(* Logix 5000 project; controller NWGG 1756-L72 rev 35.12; software revision 35.00; part 10 of 19 *)
(* tags used below, declared in another part *)
   _11_GATE_PO : ALIAS FOR I16[0];
   _123_COMPUW : ALIAS FOR I18[7];
   _12_GATE_PO : ALIAS FOR I16[1];
   _13_GATE_PO : ALIAS FOR I16[2];
   _14_GATE_PO : ALIAS FOR I16[3];
   _15_GATE_PO : ALIAS FOR I16[4];
   _16_GATE_PO : ALIAS FOR I16[5];
   _17_GATE_PO : ALIAS FOR I16[6];
   _21_GATE_PO : ALIAS FOR I16[7];
   _22_GATE_PO : ALIAS FOR I17[0];
   _23_GATE_PO : ALIAS FOR I17[1];
   _24_GATE_PO : ALIAS FOR I17[2];
   _25_GATE_PO : ALIAS FOR I17[3];
   _26_GATE_PO : ALIAS FOR I17[4];
   _27_GATE_PO : ALIAS FOR I17[5];
   _27_GATE_PO1 : ALIAS FOR N14[27];
   _28_GATE_PO : ALIAS FOR I17[6];
   _28_GATE_PO1 : ALIAS FOR N14[28];
   _29_GATE_PO : ALIAS FOR I17[7];
   _29_GATE_PO1 : ALIAS FOR N14[29];
   _41_GATE_PO : ALIAS FOR I18[0];
   _42_GATE_PO : ALIAS FOR I18[1];
   _701K_GATE2 : ALIAS FOR B21[11].2;
   _701K_VALVE : ALIAS FOR O13.10;
   Beta : BOOL;
   Calibration_Max : REAL;
   Cleaning_Motors : udt_Motor[100];
   cpTicketBinActive : DINT;
   cpTicketBinSet : DINT;
   Dev : DINT;
   I18 : INT[16];
   I18_002 : ALIAS FOR I18[2];
   I18_003 : ALIAS FOR I18[3];
   indexTbl : DINT;
   indexTRTTbl : DINT;
   InEUMax : REAL;
   MAIN_TIMER : ALIAS FOR T11[0];
   O11_000_Bit09 : ALIAS FOR O11.9;
   O11_000_Bit10 : ALIAS FOR O11.10;
   O11_000_Bit11 : ALIAS FOR O11.11;
   O11_000_Bit12 : ALIAS FOR O11.12;
   O11_000_Bit13 : ALIAS FOR O11.13;
   O11_000_Bit14 : ALIAS FOR O11.14;
   O12_000_Bit00 : ALIAS FOR O12.0;
   O12_000_Bit01 : ALIAS FOR O12.1;
   O12_000_Bit02 : ALIAS FOR O12.2;
   O16 : INT[12];
   O17 : INT[12];
   O18 : INT[12];
   O9_000_Bit00 : ALIAS FOR O9.0;
   SCREENINGS : ALIAS FOR I7.15;
   sendData : BOOL;
   sendData1 : BOOL;
   spBinGateRates : DINT[50];
   spCapGrossWt : BOOL;
   spCapTareWt : BOOL;
   spCreateTicket : BOOL;
   spShowCreateTicketPB : BOOL;
   spTicketBinActive : DINT;
   spTicketBinSet : DINT;
   spTicketProcessing : BOOL;
   spTicketProcessStr : BOOL;
   spTicketTableBay1GrsWt : DINT;
   spTicketTableBay1Wt : DINT;
   spVAR_BINARRAY : STRING[50];
   sqlIndex : DINT;
   sqlIndex1 : DINT;
   sqlNewTreatment : BOOL;
   sqlNewTreatments_ONS : DINT;
   sqlNewVariety : BOOL;
   sqlNewVariety_ONS : DINT;
   sqlTreatID : DINT;
   sqlTreatmentsRevd : DINT;
   sqlTreatRate : DINT;
   sqlTrtSendDelayTMR : TIMER;
   sqlVaritiesRevd : DINT;
   sqlVarityID : DINT;
   sqlVarityRate : DINT;
   sqlVarSendDelayTMR : TIMER;
   SWW_Index : DINT;
   SWW_Variety_DB : Varieties_DB[100];
   T11_AUTO_M : ALIAS FOR B3[11].1;
   T11_AUTO_S : ALIAS FOR B3[11].14;
   T11_SET_LO : ALIAS FOR B3[11].13;
   T12_AUTO_M : ALIAS FOR B3[12].1;
   T12_AUTO_S : ALIAS FOR B3[12].14;
   T12_SET_LO : ALIAS FOR B3[12].13;
   T13_AUTO_M : ALIAS FOR B3[13].1;
   T13_AUTO_S : ALIAS FOR B3[13].14;
   T13_SET_LO : ALIAS FOR B3[13].13;
   T14_AUTO_M : ALIAS FOR B3[14].1;
   T14_AUTO_S : ALIAS FOR B3[14].14;
   T14_SET_LO : ALIAS FOR B3[14].13;
   T15_AUTO_M : ALIAS FOR B3[15].1;
   T15_AUTO_S : ALIAS FOR B3[15].14;
   T15_SET_LO : ALIAS FOR B3[15].13;
   T16_AUTO_M : ALIAS FOR B3[16].1;
   T16_AUTO_S : ALIAS FOR B3[16].14;
   T16_SET_LO : ALIAS FOR B3[16].13;
   T17_AUTO_M : ALIAS FOR B3[17].1;
   T17_AUTO_S : ALIAS FOR B3[17].14;
   T17_SET_LO : ALIAS FOR B3[17].13;
   T21_AUTO_M : ALIAS FOR B3[21].1;
   T21_AUTO_S : ALIAS FOR B3[21].14;
   T21_SET_LO : ALIAS FOR B3[21].13;
   T22_AUTO_M : ALIAS FOR B3[22].1;
   T22_AUTO_S : ALIAS FOR B3[22].14;
   T22_SET_LO : ALIAS FOR B3[22].13;
   T23_AUTO_M : ALIAS FOR B3[23].1;
   T23_AUTO_S : ALIAS FOR B3[23].14;
   T23_SET_LO : ALIAS FOR B3[23].13;
   T24_AUTO_M : ALIAS FOR B3[24].1;
   T24_AUTO_S : ALIAS FOR B3[24].14;
   T24_SET_LO : ALIAS FOR B3[24].13;
   T25_AUTO_M : ALIAS FOR B3[25].1;
   T25_AUTO_S : ALIAS FOR B3[25].14;
   T25_SET_LO : ALIAS FOR B3[25].13;
   T26_AUTO_M : ALIAS FOR B3[26].1;
   T26_AUTO_S : ALIAS FOR B3[26].14;
   T26_SET_LO : ALIAS FOR B3[26].13;
   T27_AUTO_M : ALIAS FOR B3[27].1;
   T27_CLOSE1 : ALIAS FOR B3[27].9;
   T27_CLOSE2 : ALIAS FOR B3[27].11;
   T27_FAULT : ALIAS FOR B3[27].15;
   T27_GATE_C : ALIAS FOR C5[27];
   T27_HOLD_A : ALIAS FOR B3[27].3;
   T27_HOLD_M : ALIAS FOR B3[27].6;
   T27_OPEN_A : ALIAS FOR B3[27].8;
   T27_OPEN_M1 : ALIAS FOR B3[27].10;
   T27_RELEAS : ALIAS FOR B3[27].5;
   T27_RESET : ALIAS FOR B3[27].7;
   T27_SET_AU : ALIAS FOR B3[27].2;
   T27_STOP_A : ALIAS FOR B3[27].4;
   T28_AUTO_M : ALIAS FOR B3[28].1;
   T28_CLOSE1 : ALIAS FOR B3[28].9;
   T28_CLOSE2 : ALIAS FOR B3[28].11;
   T28_FAULT : ALIAS FOR B3[28].15;
   T28_GATE_C : ALIAS FOR C5[28];
   T28_HOLD_A : ALIAS FOR B3[28].3;
   T28_HOLD_M : ALIAS FOR B3[28].6;
   T28_OPEN_A : ALIAS FOR B3[28].8;
   T28_OPEN_M1 : ALIAS FOR B3[28].10;
   T28_RELEAS : ALIAS FOR B3[28].5;
   T28_RESET : ALIAS FOR B3[28].7;
   T28_SET_AU : ALIAS FOR B3[28].2;
   T28_STOP_A : ALIAS FOR B3[28].4;
   T29_AUTO_M : ALIAS FOR B3[29].1;
   T29_CLOSE1 : ALIAS FOR B3[29].9;
   T29_CLOSE2 : ALIAS FOR B3[29].11;
   T29_FAULT : ALIAS FOR B3[29].15;
   T29_GATE_C : ALIAS FOR C5[29];
   T29_HOLD_A : ALIAS FOR B3[29].3;
   T29_HOLD_M : ALIAS FOR B3[29].6;
   T29_OPEN_A : ALIAS FOR B3[29].8;
   T29_OPEN_M1 : ALIAS FOR B3[29].10;
   T29_RELEAS : ALIAS FOR B3[29].5;
   T29_RESET : ALIAS FOR B3[29].7;
   T29_SET_AU : ALIAS FOR B3[29].2;
   T29_STOP_A : ALIAS FOR B3[29].4;
   TestTag : REAL;
   TicketTreatPumpActive : DINT;
   TicketTreatPumpSet : DINT;
   tpCreateTicket : BOOL;
   tpCreateTicketRecvd : DINT;
   tpLocation : DINT;
   tpNewGrossWt : BOOL;
   tpNewGrossWtRecvd : DINT;
   tpNewGrossWtSent : BOOL;
   tpNewTareWt : BOOL;
   tpNewTareWtRecvd : DINT;
   tpNewTareWtSent : BOOL;
   tpShowGrossPB : BOOL;
   tpShowTarePB : BOOL;
   tpVarsTrtsComplete : BOOL;
   TRT_CNT : DINT;
   Trt_CntStore : DINT;
   TRT_TickettableItemNo : DINT[50];
   TRT_TICKETtableRate : DINT[100];
   VAR_CNT : DINT;
   VAR_CNT_ONS : DINT;
   Var_CntStore : DINT;
   VAR_TICKETtable : STRING[20];
   VAR_TickettableItemNo : DINT[50];
   VAR_TICKETtableRate : DINT[100];
   VarTrimTemp : STRING;
   zzztmpTANKtest : DINT[10];
   zzzzTestGrossWt : BOOL;
   zzzzTestTareWt : BOOL;
(* _2_MAIN, continued *)

ROUTINE _701_KValve   (* ladder *)
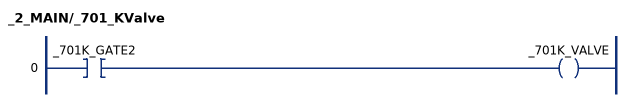
   0: XIC(_701K_GATE2)OTE(_701K_VALVE);
END_ROUTINE

ROUTINE _99_Scaling   (* function block diagram *)
   SHEET 1
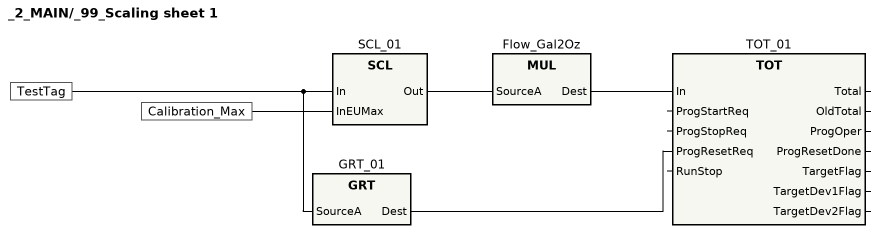
   GRT_01 : GRT(SourceA := TestTag);
   SCL_01 : SCL(In := TestTag, InEUMax := Calibration_Max);
   Flow_Gal2Oz : MUL(SourceA := SCL_01.Out);
   TOT_01 : TOT(In := Flow_Gal2Oz.Dest, ProgResetReq := GRT_01.Dest);   // unwired pins: ProgStartReq ProgStopReq Total OldTotal ProgOper RunStop ProgResetDone TargetFlag TargetDev1Flag TargetDev2Flag
   SHEET 2
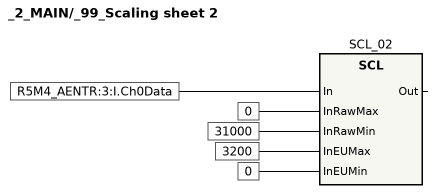
   SCL_02 : SCL(In := R5M4_AENTR:3:I.Ch0Data, InRawMax := 0, InRawMin := 31000, InEUMax := 3200, InEUMin := 0);   // unwired pins: Out
END_ROUTINE
END_PROGRAM

PROGRAM Amp_Guages   (* main routine Amp_Guages *)
VAR
   SCL_AMP_Belt11 : SCALE := (In := 28.19336, InRawMax := 6000.0, InEUMax := 1.61, Out := 0.007565218);
   SCL_AMP_Belt11_01 : SCALE := (In := 23.047852, InRawMax := 9000.0, InRawMin := 20.0, InEUMax := 2.15, Out := 0.0007297195);
   SCL_AMP_Belt11_02 : SCALE := (In := 4111.1504, InRawMax := 7000.0, InRawMin := 20.0, InEUMax := 1.61, Out := 0.94366074);
   SCL_AMP_Belt11_03 : SCALE := (In := 7592.727, InRawMax := 13000.0, InRawMin := 20.0, InEUMax := 3.88, Out := 2.2636504);
END_VAR

ROUTINE Amp_Guages   (* function block diagram *)
   SHEET 1
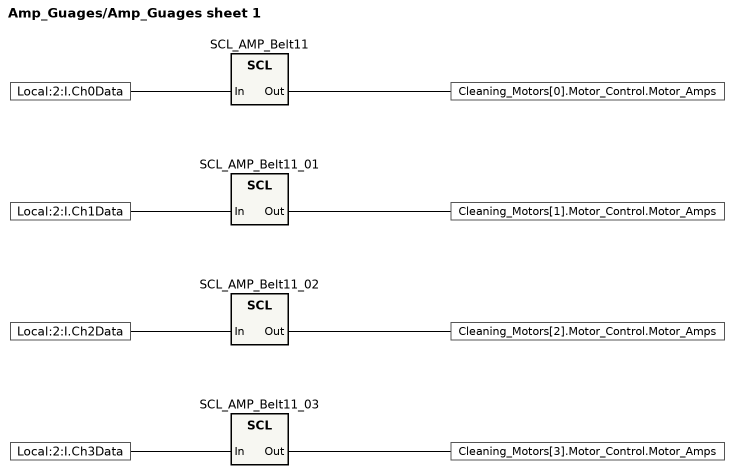
   SCL_AMP_Belt11 : SCL(In := Local:2:I.Ch0Data);
   SCL_AMP_Belt11_01 : SCL(In := Local:2:I.Ch1Data);
   SCL_AMP_Belt11_02 : SCL(In := Local:2:I.Ch2Data);
   SCL_AMP_Belt11_03 : SCL(In := Local:2:I.Ch3Data);
   Cleaning_Motors[0].Motor_Control.Motor_Amps := SCL_AMP_Belt11.Out;
   Cleaning_Motors[1].Motor_Control.Motor_Amps := SCL_AMP_Belt11_01.Out;
   Cleaning_Motors[2].Motor_Control.Motor_Amps := SCL_AMP_Belt11_02.Out;
   Cleaning_Motors[3].Motor_Control.Motor_Amps := SCL_AMP_Belt11_03.Out;
END_ROUTINE
END_PROGRAM

PROGRAM Load_Requests   (* main routine Main *)

ROUTINE Main   (* ladder *)
END_ROUTINE
END_PROGRAM

PROGRAM Main   (* main routine Main *)
VAR
   alm_Development : ALARM_DIGITAL;
   Beta_Mode : BOOL;
END_VAR

ROUTINE Main   (* ladder *)
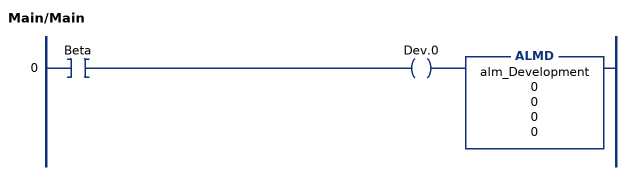
   0: XIC(Beta)OTE(Dev.0)ALMD(alm_Development,0,0,0,0);
END_ROUTINE
END_PROGRAM

PROGRAM MainProgram   (* main routine MainRoutine *)
VAR
   Alm_Test : BOOL := 1;
   ATestAck : BOOL;
   ATestPDis : BOOL;
   ATestPEna : BOOL;
   ATestReset : BOOL;
   BIN13test : BOOL;
   CleaningBinVarieties : STRING[10] := ([2] := 'hale', [3] := 'Hale full', [4] := 'Hale', [6] := 'HD307 Screenings');
   CTR_Scale_Accum_Rate_Index : COUNTER;
   Flow_Gal2Oz : FBD_MATH := (SourceA := 4000.0, SourceB := 0.25, Dest := 1000.0);
   GRT_01 : FBD_COMPARE := (SourceB := 75.0);
   Rate_Tmr : TIMER := (PRE := 1000, ACC := 610, TT := 1, DN := 1);
   Scale_Avg_Ctr : COUNTER := (PRE := 10, ACC := 2, CU := 1);
   ScaleWeights : DINT[60];
   SCL_01 : SCALE := (InRawMax := 100.0, InEUMax := 4000.0);
   SCL_02 : SCALE := (In := 16384.0, InRawMax := 13975.0, InRawMin := 578.0, InEUMax := 3000.0, Limiting := 1, Out := 3000.0, MaxAlarm := 1);
   Tare : DINT;
   tmr_User_Cancel : TIMER := (PRE := 5000, ACC := 5004, EN := 1, DN := 1);
   tmrWeightTest : TIMER := (PRE := 500, ACC := 112, EN := 1, TT := 1);
   TOT_01 : TOTALIZER := (TimeBase := 1, Gain := 1.0, ProgProgReq := 1, ProgStartReq := 1, ProgStopReq := 1, RTSTime := 1, Total := 4074.4673, OldTotal := 9541.935, ProgOper := 1, TargetFlag := 1, TargetDev1Flag := 1, TargetDev2Flag := 1, LowInCutoffFlag := 1, DeltaT := 0.016);
   Truck_Scale_Control : Truck_Scale_Control[2];
   Weight_Seed : DINT := 10;
END_VAR

ROUTINE _100_VarCfg   (* ladder *)
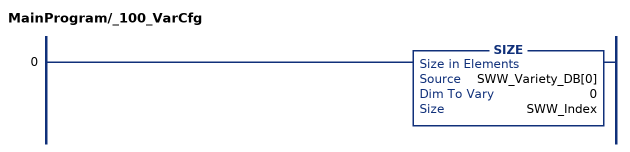
   0: SIZE(SWW_Variety_DB[0],0,SWW_Index);
END_ROUTINE

ROUTINE _31_TANK_27   (* ladder *)
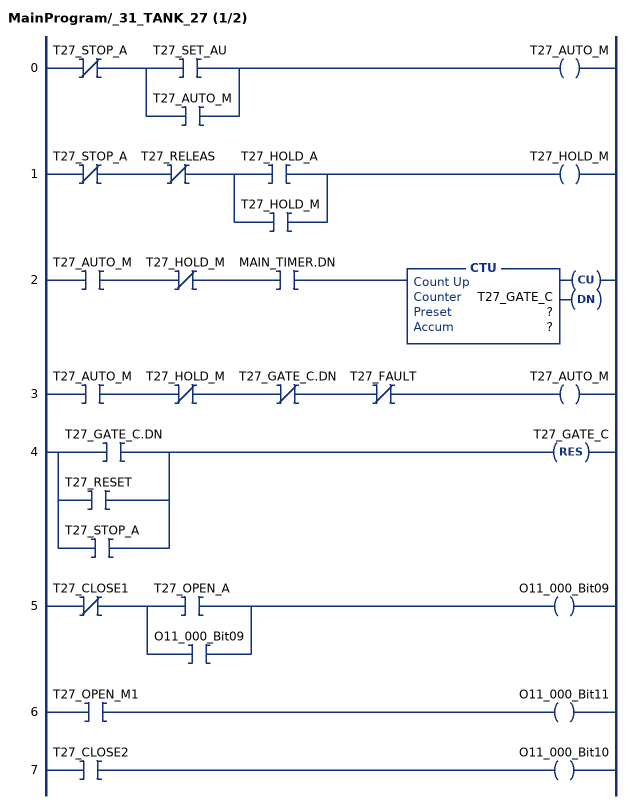
   0: XIO(T27_STOP_A)[XIC(T27_SET_AU) ,XIC(T27_AUTO_M) ]OTE(T27_AUTO_M);
   1: XIO(T27_STOP_A)XIO(T27_RELEAS)[XIC(T27_HOLD_A) ,XIC(T27_HOLD_M) ]OTE(T27_HOLD_M);
   2: XIC(T27_AUTO_M)XIO(T27_HOLD_M)XIC(MAIN_TIMER.DN)CTU(T27_GATE_C,?,?);
   3: XIC(T27_AUTO_M)XIO(T27_HOLD_M)XIO(T27_GATE_C.DN)XIO(T27_FAULT)OTE(T27_AUTO_M);
   4: [XIC(T27_GATE_C.DN) ,XIC(T27_RESET) ,XIC(T27_STOP_A) ]RES(T27_GATE_C);
   5: XIO(T27_CLOSE1)[XIC(T27_OPEN_A) ,XIC(O11_000_Bit09) ]OTE(O11_000_Bit09);
   6: XIC(T27_OPEN_M1)OTE(O11_000_Bit11);
   7: XIC(T27_CLOSE2)OTE(O11_000_Bit10);
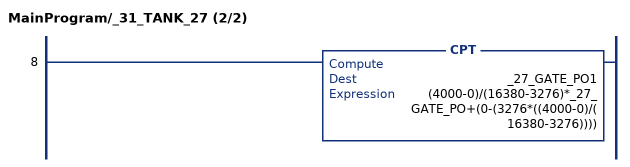
   8: CPT(_27_GATE_PO1,(4000-0)/(16380-3276)*_27_GATE_PO+(0-(3276*((4000-0)/(16380-3276)))));
END_ROUTINE

ROUTINE _32_TANK_28   (* ladder *)
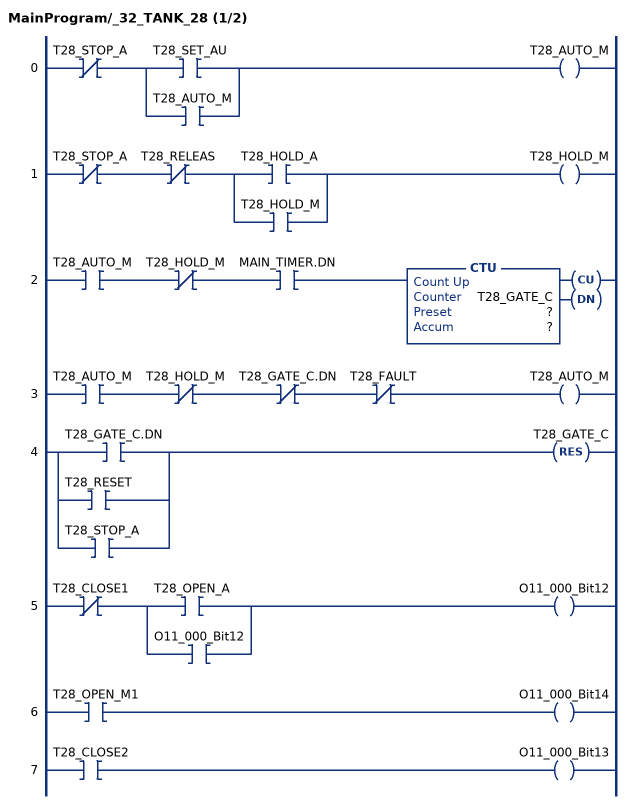
   0: XIO(T28_STOP_A)[XIC(T28_SET_AU) ,XIC(T28_AUTO_M) ]OTE(T28_AUTO_M);
   1: XIO(T28_STOP_A)XIO(T28_RELEAS)[XIC(T28_HOLD_A) ,XIC(T28_HOLD_M) ]OTE(T28_HOLD_M);
   2: XIC(T28_AUTO_M)XIO(T28_HOLD_M)XIC(MAIN_TIMER.DN)CTU(T28_GATE_C,?,?);
   3: XIC(T28_AUTO_M)XIO(T28_HOLD_M)XIO(T28_GATE_C.DN)XIO(T28_FAULT)OTE(T28_AUTO_M);
   4: [XIC(T28_GATE_C.DN) ,XIC(T28_RESET) ,XIC(T28_STOP_A) ]RES(T28_GATE_C);
   5: XIO(T28_CLOSE1)[XIC(T28_OPEN_A) ,XIC(O11_000_Bit12) ]OTE(O11_000_Bit12);
   6: XIC(T28_OPEN_M1)OTE(O11_000_Bit14);
   7: XIC(T28_CLOSE2)OTE(O11_000_Bit13);
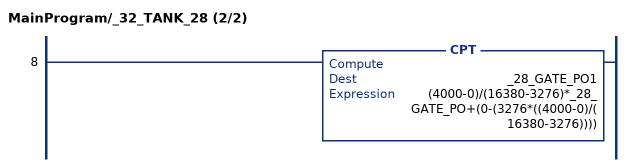
   8: CPT(_28_GATE_PO1,(4000-0)/(16380-3276)*_28_GATE_PO+(0-(3276*((4000-0)/(16380-3276)))));
END_ROUTINE

ROUTINE _33_TANK_29   (* ladder *)
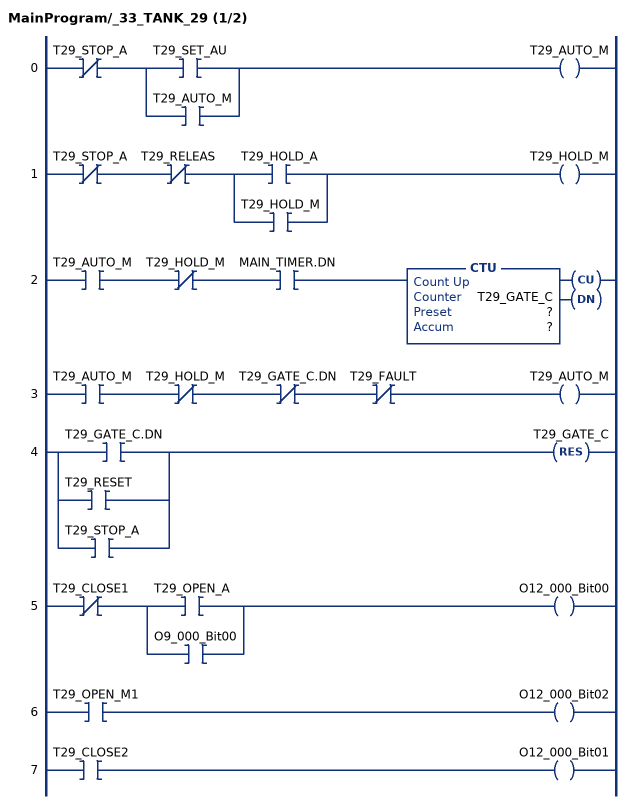
   0: XIO(T29_STOP_A)[XIC(T29_SET_AU) ,XIC(T29_AUTO_M) ]OTE(T29_AUTO_M);
   1: XIO(T29_STOP_A)XIO(T29_RELEAS)[XIC(T29_HOLD_A) ,XIC(T29_HOLD_M) ]OTE(T29_HOLD_M);
   2: XIC(T29_AUTO_M)XIO(T29_HOLD_M)XIC(MAIN_TIMER.DN)CTU(T29_GATE_C,?,?);
   3: XIC(T29_AUTO_M)XIO(T29_HOLD_M)XIO(T29_GATE_C.DN)XIO(T29_FAULT)OTE(T29_AUTO_M);
   4: [XIC(T29_GATE_C.DN) ,XIC(T29_RESET) ,XIC(T29_STOP_A) ]RES(T29_GATE_C);
   5: XIO(T29_CLOSE1)[XIC(T29_OPEN_A) ,XIC(O9_000_Bit00) ]OTE(O12_000_Bit00);
   6: XIC(T29_OPEN_M1)OTE(O12_000_Bit02);
   7: XIC(T29_CLOSE2)OTE(O12_000_Bit01);
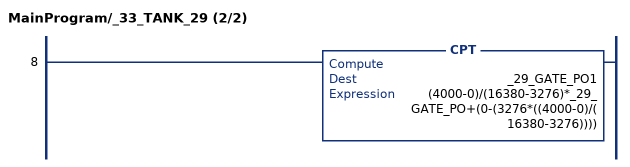
   8: CPT(_29_GATE_PO1,(4000-0)/(16380-3276)*_29_GATE_PO+(0-(3276*((4000-0)/(16380-3276)))));
END_ROUTINE

ROUTINE ANALOG_SCALING   (* ladder *)
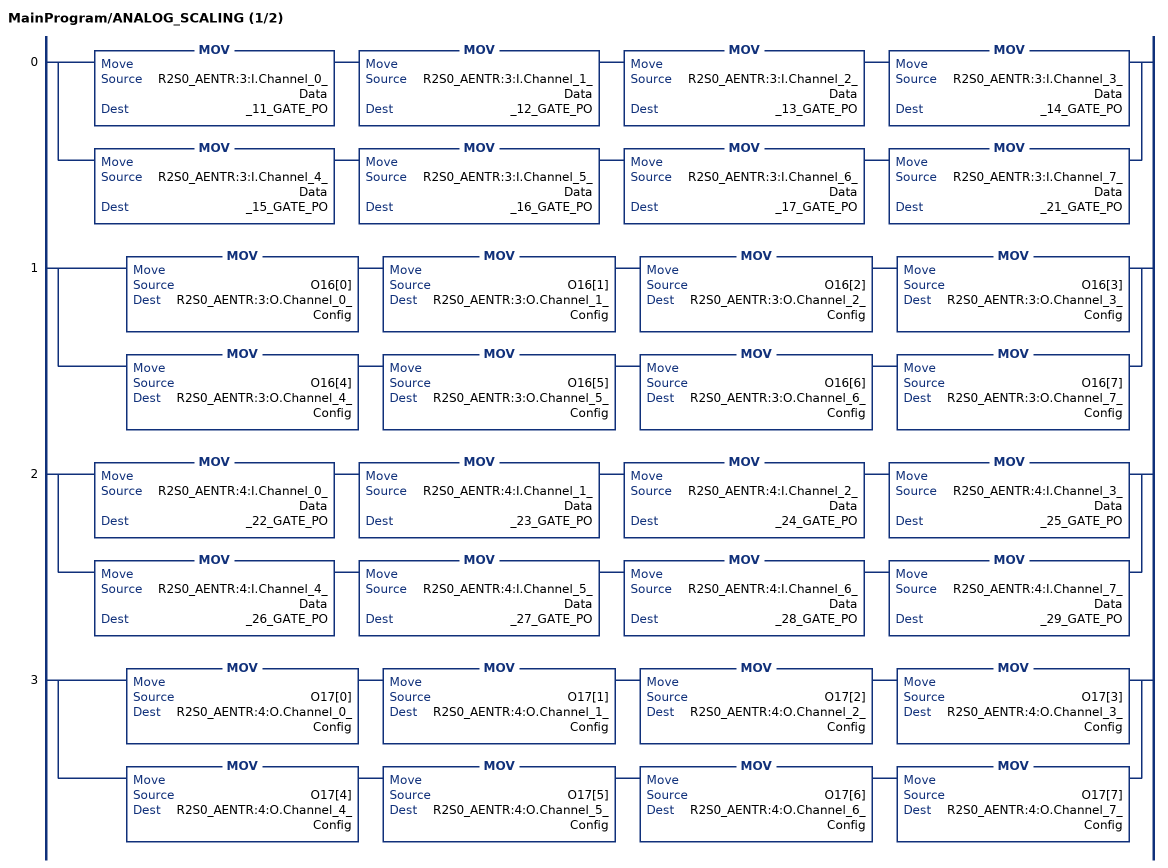
   0: [MOV(R2S0_AENTR:3:I.Channel_0_Data,_11_GATE_PO) MOV(R2S0_AENTR:3:I.Channel_1_Data,_12_GATE_PO) MOV(R2S0_AENTR:3:I.Channel_2_Data,_13_GATE_PO) MOV(R2S0_AENTR:3:I.Channel_3_Data,_14_GATE_PO) ,MOV(R2S0_AENTR:3:I.Channel_4_Data,_15_GATE_PO) MOV(R2S0_AENTR:3:I.Channel_5_Data,_16_GATE_PO) MOV(R2S0_AENTR:3:I.Channel_6_Data,_17_GATE_PO) MOV(R2S0_AENTR:3:I.Channel_7_Data,_21_GATE_PO) ];
   1: [MOV(O16[0],R2S0_AENTR:3:O.Channel_0_Config) MOV(O16[1],R2S0_AENTR:3:O.Channel_1_Config) MOV(O16[2],R2S0_AENTR:3:O.Channel_2_Config) MOV(O16[3],R2S0_AENTR:3:O.Channel_3_Config) ,MOV(O16[4],R2S0_AENTR:3:O.Channel_4_Config) MOV(O16[5],R2S0_AENTR:3:O.Channel_5_Config) MOV(O16[6],R2S0_AENTR:3:O.Channel_6_Config) MOV(O16[7],R2S0_AENTR:3:O.Channel_7_Config) ];
   2: [MOV(R2S0_AENTR:4:I.Channel_0_Data,_22_GATE_PO) MOV(R2S0_AENTR:4:I.Channel_1_Data,_23_GATE_PO) MOV(R2S0_AENTR:4:I.Channel_2_Data,_24_GATE_PO) MOV(R2S0_AENTR:4:I.Channel_3_Data,_25_GATE_PO) ,MOV(R2S0_AENTR:4:I.Channel_4_Data,_26_GATE_PO) MOV(R2S0_AENTR:4:I.Channel_5_Data,_27_GATE_PO) MOV(R2S0_AENTR:4:I.Channel_6_Data,_28_GATE_PO) MOV(R2S0_AENTR:4:I.Channel_7_Data,_29_GATE_PO) ];
   3: [MOV(O17[0],R2S0_AENTR:4:O.Channel_0_Config) MOV(O17[1],R2S0_AENTR:4:O.Channel_1_Config) MOV(O17[2],R2S0_AENTR:4:O.Channel_2_Config) MOV(O17[3],R2S0_AENTR:4:O.Channel_3_Config) ,MOV(O17[4],R2S0_AENTR:4:O.Channel_4_Config) MOV(O17[5],R2S0_AENTR:4:O.Channel_5_Config) MOV(O17[6],R2S0_AENTR:4:O.Channel_6_Config) MOV(O17[7],R2S0_AENTR:4:O.Channel_7_Config) ];
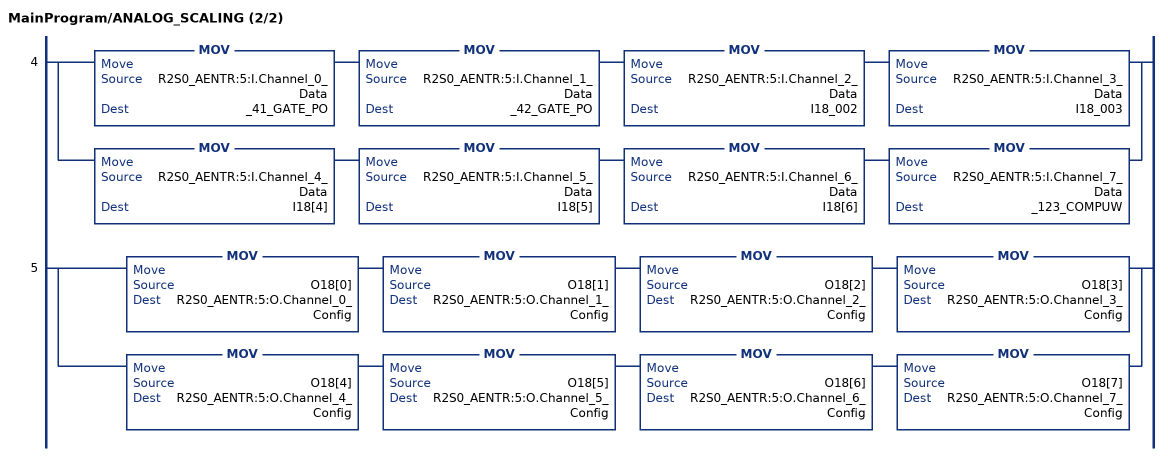
   4: [MOV(R2S0_AENTR:5:I.Channel_0_Data,_41_GATE_PO) MOV(R2S0_AENTR:5:I.Channel_1_Data,_42_GATE_PO) MOV(R2S0_AENTR:5:I.Channel_2_Data,I18_002) MOV(R2S0_AENTR:5:I.Channel_3_Data,I18_003) ,MOV(R2S0_AENTR:5:I.Channel_4_Data,I18[4]) MOV(R2S0_AENTR:5:I.Channel_5_Data,I18[5]) MOV(R2S0_AENTR:5:I.Channel_6_Data,I18[6]) MOV(R2S0_AENTR:5:I.Channel_7_Data,_123_COMPUW) ];
   5: [MOV(O18[0],R2S0_AENTR:5:O.Channel_0_Config) MOV(O18[1],R2S0_AENTR:5:O.Channel_1_Config) MOV(O18[2],R2S0_AENTR:5:O.Channel_2_Config) MOV(O18[3],R2S0_AENTR:5:O.Channel_3_Config) ,MOV(O18[4],R2S0_AENTR:5:O.Channel_4_Config) MOV(O18[5],R2S0_AENTR:5:O.Channel_5_Config) MOV(O18[6],R2S0_AENTR:5:O.Channel_6_Config) MOV(O18[7],R2S0_AENTR:5:O.Channel_7_Config) ];
END_ROUTINE

ROUTINE DATA   (* ladder *)
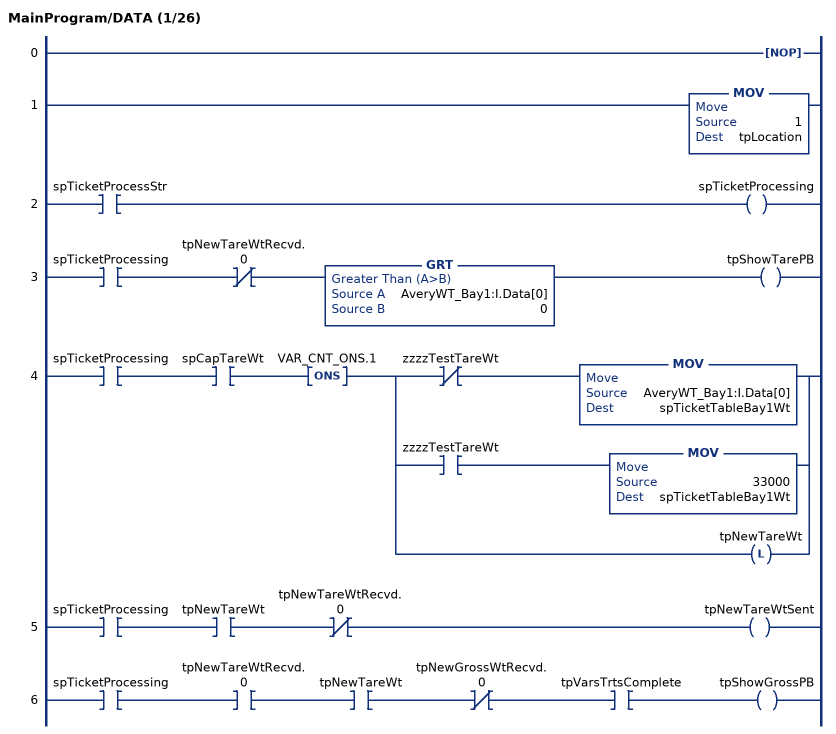
   0: NOP();
   1: MOV(1,tpLocation);
   2: XIC(spTicketProcessStr)OTE(spTicketProcessing);
   3: XIC(spTicketProcessing)XIO(tpNewTareWtRecvd.0)GRT(AveryWT_Bay1:I.Data[0],0)OTE(tpShowTarePB);
   4: XIC(spTicketProcessing)XIC(spCapTareWt)ONS(VAR_CNT_ONS.1)[XIO(zzzzTestTareWt) MOV(AveryWT_Bay1:I.Data[0],spTicketTableBay1Wt) ,XIC(zzzzTestTareWt) MOV(33000,spTicketTableBay1Wt) ,OTL(tpNewTareWt) ];
   5: XIC(spTicketProcessing)XIC(tpNewTareWt)XIO(tpNewTareWtRecvd.0)OTE(tpNewTareWtSent);
   6: XIC(spTicketProcessing)XIC(tpNewTareWtRecvd.0)XIC(tpNewTareWt)XIO(tpNewGrossWtRecvd.0)XIC(tpVarsTrtsComplete)OTE(tpShowGrossPB);
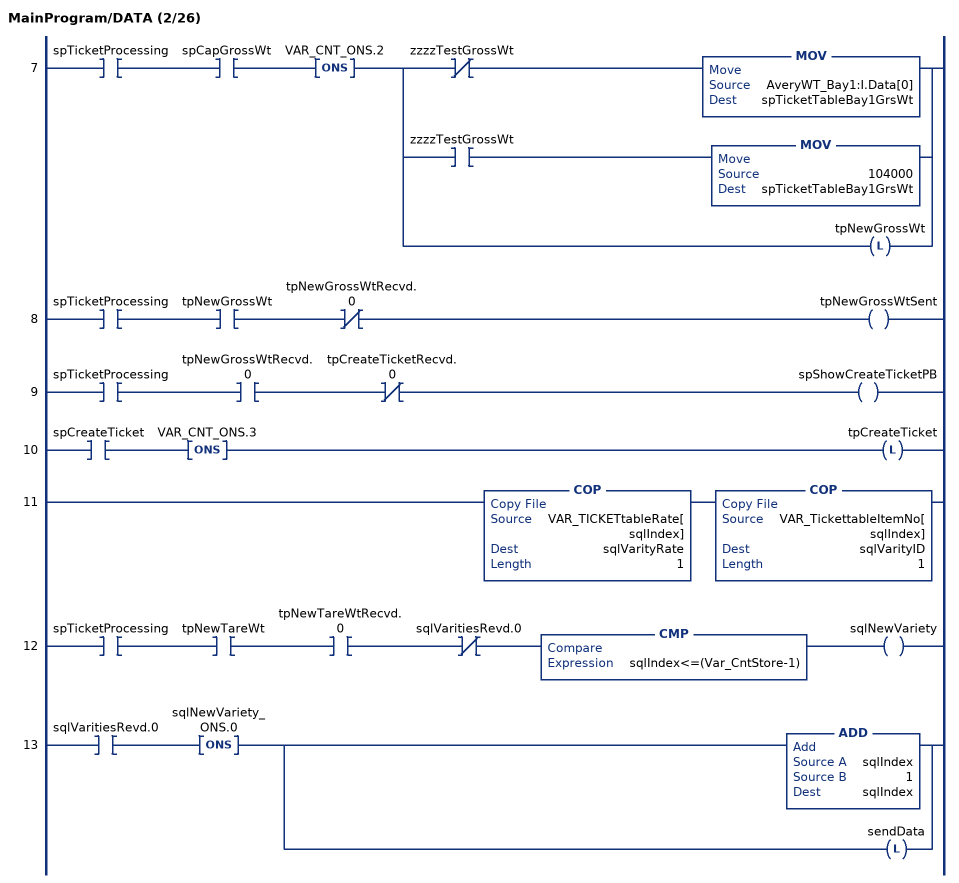
   7: XIC(spTicketProcessing)XIC(spCapGrossWt)ONS(VAR_CNT_ONS.2)[XIO(zzzzTestGrossWt) MOV(AveryWT_Bay1:I.Data[0],spTicketTableBay1GrsWt) ,XIC(zzzzTestGrossWt) MOV(104000,spTicketTableBay1GrsWt) ,OTL(tpNewGrossWt) ];
   8: XIC(spTicketProcessing)XIC(tpNewGrossWt)XIO(tpNewGrossWtRecvd.0)OTE(tpNewGrossWtSent);
   9: XIC(spTicketProcessing)XIC(tpNewGrossWtRecvd.0)XIO(tpCreateTicketRecvd.0)OTE(spShowCreateTicketPB);
   10: XIC(spCreateTicket)ONS(VAR_CNT_ONS.3)OTL(tpCreateTicket);
   11: COP(VAR_TICKETtableRate[sqlIndex],sqlVarityRate,1)COP(VAR_TickettableItemNo[sqlIndex],sqlVarityID,1);
   12: XIC(spTicketProcessing)XIC(tpNewTareWt)XIC(tpNewTareWtRecvd.0)XIO(sqlVaritiesRevd.0)CMP(sqlIndex<=(Var_CntStore-1))OTE(sqlNewVariety);
   13: XIC(sqlVaritiesRevd.0)ONS(sqlNewVariety_ONS.0)[ADD(sqlIndex,1,sqlIndex) ,OTL(sendData) ];
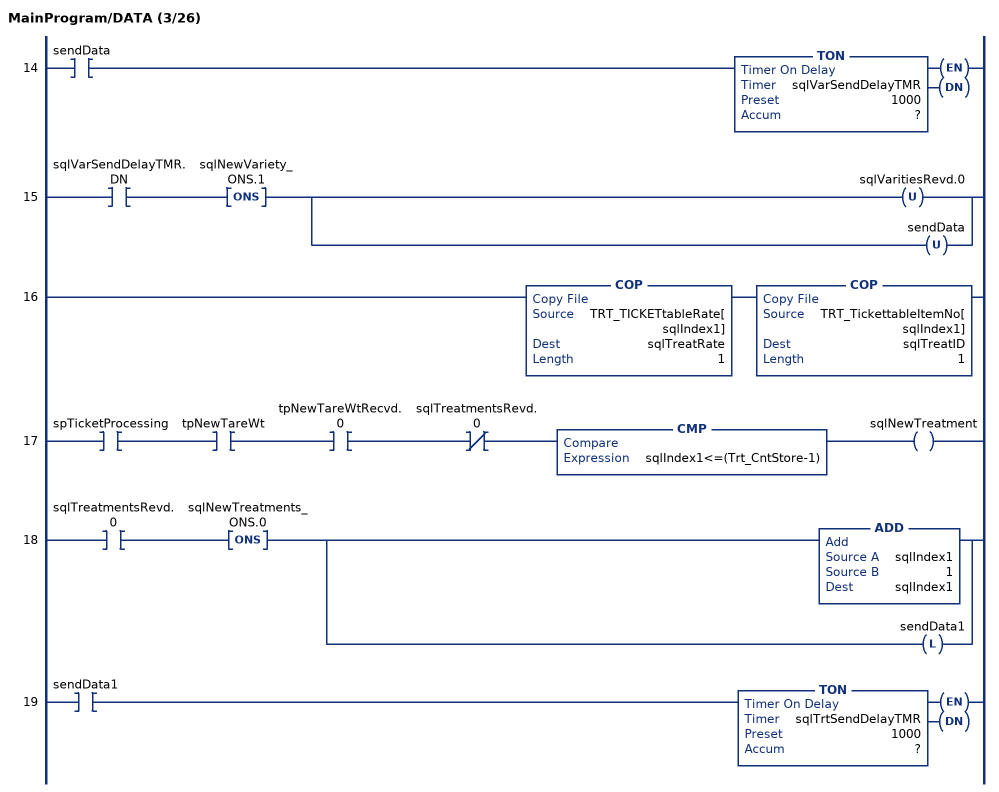
   14: XIC(sendData)TON(sqlVarSendDelayTMR,?,?);
   15: XIC(sqlVarSendDelayTMR.DN)ONS(sqlNewVariety_ONS.1)[OTU(sqlVaritiesRevd.0) ,OTU(sendData) ];
   16: COP(TRT_TICKETtableRate[sqlIndex1],sqlTreatRate,1)COP(TRT_TickettableItemNo[sqlIndex1],sqlTreatID,1);
   17: XIC(spTicketProcessing)XIC(tpNewTareWt)XIC(tpNewTareWtRecvd.0)XIO(sqlTreatmentsRevd.0)CMP(sqlIndex1<=(Trt_CntStore-1))OTE(sqlNewTreatment);
   18: XIC(sqlTreatmentsRevd.0)ONS(sqlNewTreatments_ONS.0)[ADD(sqlIndex1,1,sqlIndex1) ,OTL(sendData1) ];
   19: XIC(sendData1)TON(sqlTrtSendDelayTMR,?,?);
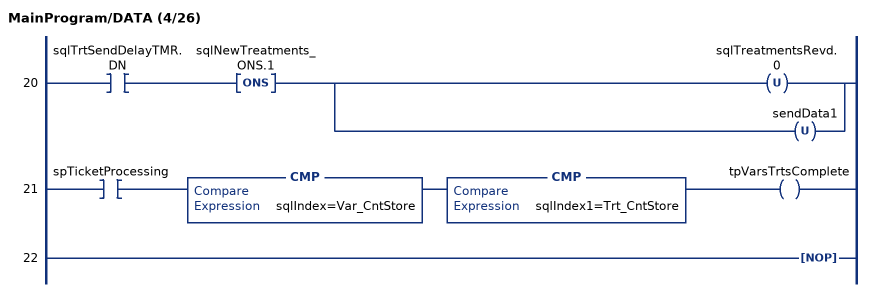
   20: XIC(sqlTrtSendDelayTMR.DN)ONS(sqlNewTreatments_ONS.1)[OTU(sqlTreatmentsRevd.0) ,OTU(sendData1) ];
   21: XIC(spTicketProcessing)CMP(sqlIndex=Var_CntStore)CMP(sqlIndex1=Trt_CntStore)OTE(tpVarsTrtsComplete);
   22: NOP();
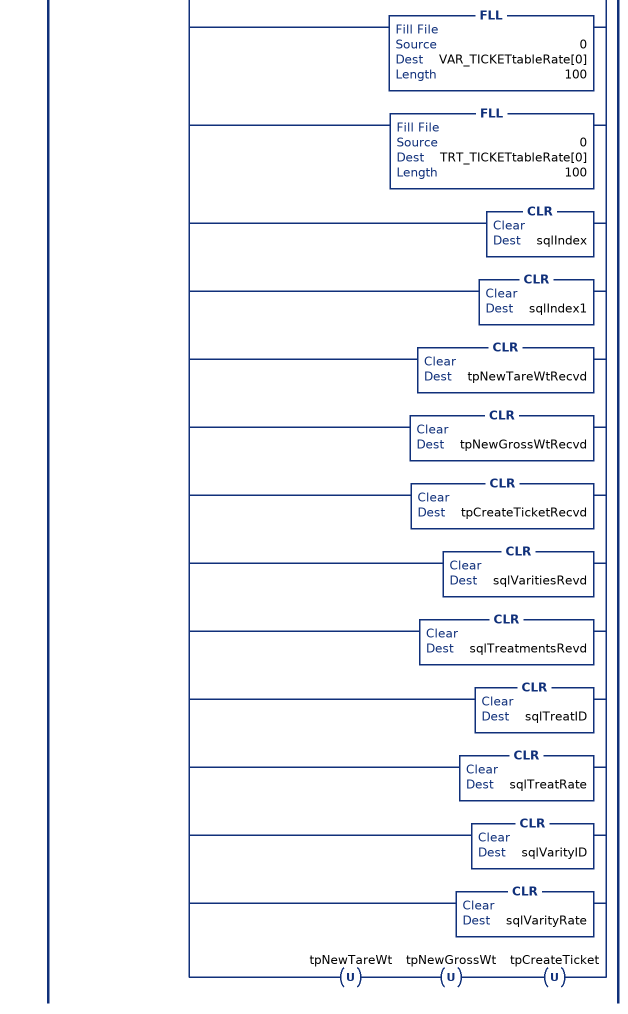
   23: XIO(spTicketProcessing)[CLR(VAR_CNT) ,CLR(cpTicketBinActive) ,CLR(spTicketBinActive) ,CLR(cpTicketBinSet) ,CLR(spTicketBinSet) ,CLR(indexTbl) ,CLR(indexTRTTbl) ,CLR(TRT_CNT) ,CLR(TicketTreatPumpActive) ,CLR(TicketTreatPumpSet) ,CLR(spTicketTableBay1Wt) ,CLR(spTicketTableBay1GrsWt) ,FLL(0,VAR_TickettableItemNo[0],50) ,FLL(0,TRT_TickettableItemNo[0],50) ,FLL(0,VAR_TICKETtableRate[0],100) ,FLL(0,TRT_TICKETtableRate[0],100) ,CLR(sqlIndex) ,CLR(sqlIndex1) ,CLR(tpNewTareWtRecvd) ,CLR(tpNewGrossWtRecvd) ,CLR(tpCreateTicketRecvd) ,CLR(sqlVaritiesRevd) ,CLR(sqlTreatmentsRevd) ,CLR(sqlTreatID) ,CLR(sqlTreatRate) ,CLR(sqlVarityID) ,CLR(sqlVarityRate) ,OTU(tpNewTareWt) OTU(tpNewGrossWt) OTU(tpCreateTicket) ];
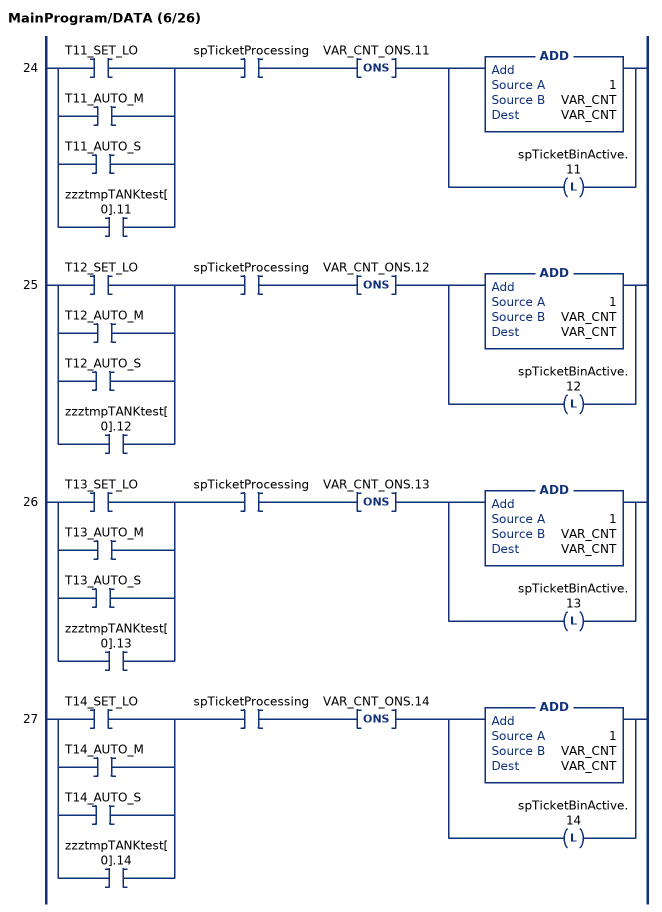
   24: [XIC(T11_SET_LO) ,XIC(T11_AUTO_M) ,XIC(T11_AUTO_S) ,XIC(zzztmpTANKtest[0].11) ]XIC(spTicketProcessing)ONS(VAR_CNT_ONS.11)[ADD(1,VAR_CNT,VAR_CNT) ,OTL(spTicketBinActive.11) ];
   25: [XIC(T12_SET_LO) ,XIC(T12_AUTO_M) ,XIC(T12_AUTO_S) ,XIC(zzztmpTANKtest[0].12) ]XIC(spTicketProcessing)ONS(VAR_CNT_ONS.12)[ADD(1,VAR_CNT,VAR_CNT) ,OTL(spTicketBinActive.12) ];
   26: [XIC(T13_SET_LO) ,XIC(T13_AUTO_M) ,XIC(T13_AUTO_S) ,XIC(zzztmpTANKtest[0].13) ]XIC(spTicketProcessing)ONS(VAR_CNT_ONS.13)[ADD(1,VAR_CNT,VAR_CNT) ,OTL(spTicketBinActive.13) ];
   27: [XIC(T14_SET_LO) ,XIC(T14_AUTO_M) ,XIC(T14_AUTO_S) ,XIC(zzztmpTANKtest[0].14) ]XIC(spTicketProcessing)ONS(VAR_CNT_ONS.14)[ADD(1,VAR_CNT,VAR_CNT) ,OTL(spTicketBinActive.14) ];
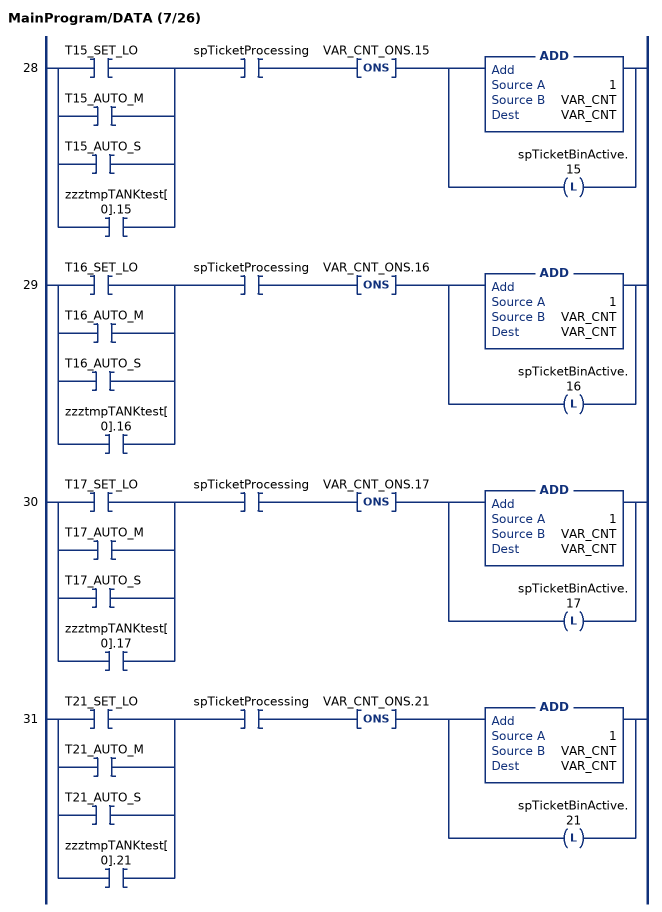
   28: [XIC(T15_SET_LO) ,XIC(T15_AUTO_M) ,XIC(T15_AUTO_S) ,XIC(zzztmpTANKtest[0].15) ]XIC(spTicketProcessing)ONS(VAR_CNT_ONS.15)[ADD(1,VAR_CNT,VAR_CNT) ,OTL(spTicketBinActive.15) ];
   29: [XIC(T16_SET_LO) ,XIC(T16_AUTO_M) ,XIC(T16_AUTO_S) ,XIC(zzztmpTANKtest[0].16) ]XIC(spTicketProcessing)ONS(VAR_CNT_ONS.16)[ADD(1,VAR_CNT,VAR_CNT) ,OTL(spTicketBinActive.16) ];
   30: [XIC(T17_SET_LO) ,XIC(T17_AUTO_M) ,XIC(T17_AUTO_S) ,XIC(zzztmpTANKtest[0].17) ]XIC(spTicketProcessing)ONS(VAR_CNT_ONS.17)[ADD(1,VAR_CNT,VAR_CNT) ,OTL(spTicketBinActive.17) ];
   31: [XIC(T21_SET_LO) ,XIC(T21_AUTO_M) ,XIC(T21_AUTO_S) ,XIC(zzztmpTANKtest[0].21) ]XIC(spTicketProcessing)ONS(VAR_CNT_ONS.21)[ADD(1,VAR_CNT,VAR_CNT) ,OTL(spTicketBinActive.21) ];
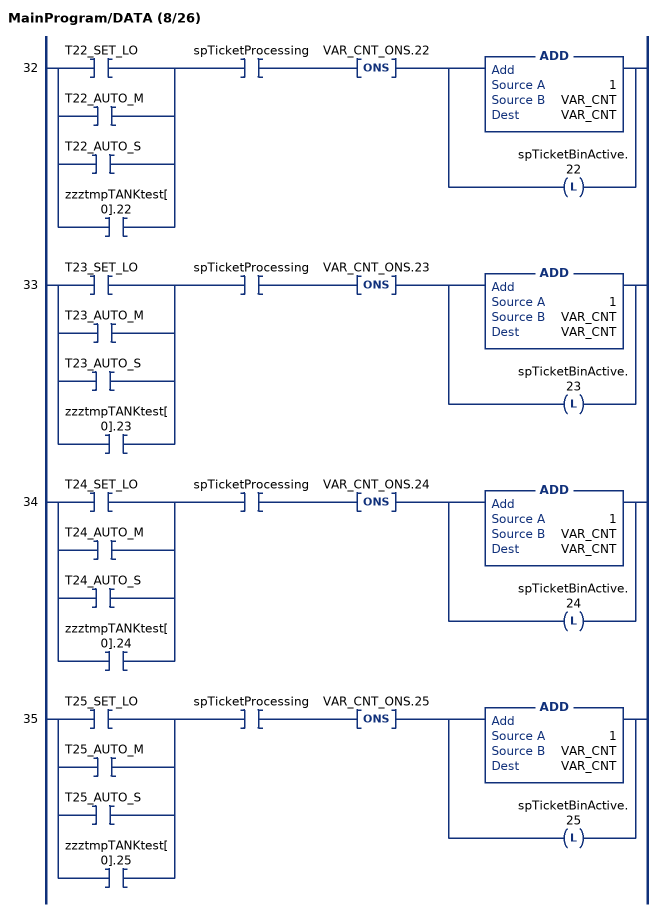
   32: [XIC(T22_SET_LO) ,XIC(T22_AUTO_M) ,XIC(T22_AUTO_S) ,XIC(zzztmpTANKtest[0].22) ]XIC(spTicketProcessing)ONS(VAR_CNT_ONS.22)[ADD(1,VAR_CNT,VAR_CNT) ,OTL(spTicketBinActive.22) ];
   33: [XIC(T23_SET_LO) ,XIC(T23_AUTO_M) ,XIC(T23_AUTO_S) ,XIC(zzztmpTANKtest[0].23) ]XIC(spTicketProcessing)ONS(VAR_CNT_ONS.23)[ADD(1,VAR_CNT,VAR_CNT) ,OTL(spTicketBinActive.23) ];
   34: [XIC(T24_SET_LO) ,XIC(T24_AUTO_M) ,XIC(T24_AUTO_S) ,XIC(zzztmpTANKtest[0].24) ]XIC(spTicketProcessing)ONS(VAR_CNT_ONS.24)[ADD(1,VAR_CNT,VAR_CNT) ,OTL(spTicketBinActive.24) ];
   35: [XIC(T25_SET_LO) ,XIC(T25_AUTO_M) ,XIC(T25_AUTO_S) ,XIC(zzztmpTANKtest[0].25) ]XIC(spTicketProcessing)ONS(VAR_CNT_ONS.25)[ADD(1,VAR_CNT,VAR_CNT) ,OTL(spTicketBinActive.25) ];
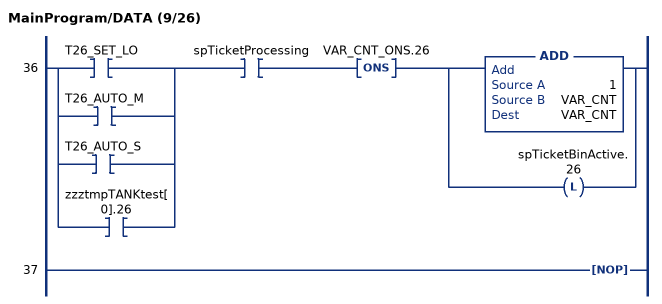
   36: [XIC(T26_SET_LO) ,XIC(T26_AUTO_M) ,XIC(T26_AUTO_S) ,XIC(zzztmpTANKtest[0].26) ]XIC(spTicketProcessing)ONS(VAR_CNT_ONS.26)[ADD(1,VAR_CNT,VAR_CNT) ,OTL(spTicketBinActive.26) ];
   37: NOP();
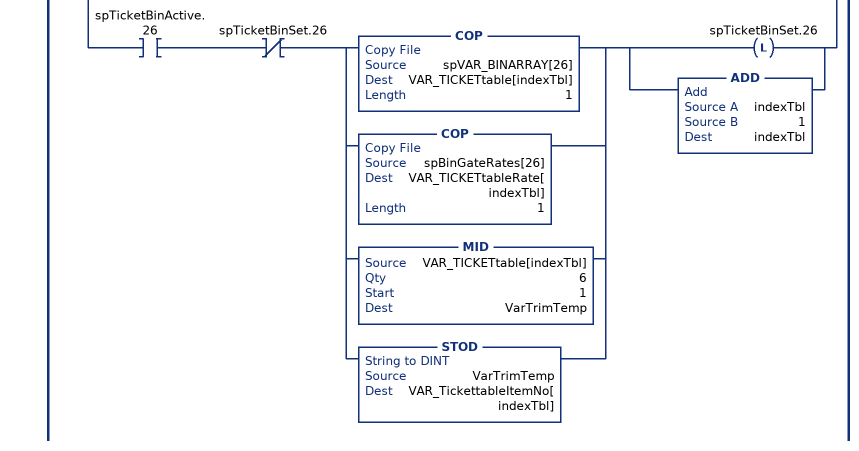
   38: GRT(VAR_CNT,0)LES(indexTbl,VAR_CNT)[XIC(spTicketBinActive.11) XIO(spTicketBinSet.11) [COP(spVAR_BINARRAY[11],VAR_TICKETtable[indexTbl],1) ,COP(spBinGateRates[11],VAR_TICKETtableRate[indexTbl],1) ,MID(VAR_TICKETtable[indexTbl],6,1,VarTrimTemp) ,STOD(VarTrimTemp,VAR_TickettableItemNo[indexTbl]) ] [OTL(spTicketBinSet.11) ,ADD(indexTbl,1,indexTbl) ] ,XIC(spTicketBinActive.12) XIO(spTicketBinSet.12) [COP(spVAR_BINARRAY[12],VAR_TICKETtable[indexTbl],1) ,COP(spBinGateRates[12],VAR_TICKETtableRate[indexTbl],1) ,MID(VAR_TICKETtable[indexTbl],6,1,VarTrimTemp) ,STOD(VarTrimTemp,VAR_TickettableItemNo[indexTbl]) ] [OTL(spTicketBinSet.12) ,ADD(indexTbl,1,indexTbl) ] ,XIC(spTicketBinActive.13) XIO(spTicketBinSet.13) [COP(spVAR_BINARRAY[13],VAR_TICKETtable[indexTbl],1) ,COP(spBinGateRates[13],VAR_TICKETtableRate[indexTbl],1) ,MID(VAR_TICKETtable[indexTbl],6,1,VarTrimTemp) ,STOD(VarTrimTemp,VAR_TickettableItemNo[indexTbl]) ] [OTL(spTicketBinSet.13) ,ADD(indexTbl,1,indexTbl) ] ,XIC(spTicketBinActive.14) XIO(spTicketBinSet.14) [COP(spVAR_BINARRAY[14],VAR_TICKETtable[indexTbl],1) ,COP(spBinGateRates[14],VAR_TICKETtableRate[indexTbl],1) ,MID(VAR_TICKETtable[indexTbl],6,1,VarTrimTemp) ,STOD(VarTrimTemp,VAR_TickettableItemNo[indexTbl]) ] [OTL(spTicketBinSet.14) ,ADD(indexTbl,1,indexTbl) ] ,XIC(spTicketBinActive.15) XIO(spTicketBinSet.15) [COP(spVAR_BINARRAY[15],VAR_TICKETtable[indexTbl],1) ,COP(spBinGateRates[15],VAR_TICKETtableRate[indexTbl],1) ,MID(VAR_TICKETtable[indexTbl],6,1,VarTrimTemp) ,STOD(VarTrimTemp,VAR_TickettableItemNo[indexTbl]) ] [OTL(spTicketBinSet.15) ,ADD(indexTbl,1,indexTbl) ] ,XIC(spTicketBinActive.16) XIO(spTicketBinSet.16) [COP(spVAR_BINARRAY[16],VAR_TICKETtable[indexTbl],1) ,COP(spBinGateRates[16],VAR_TICKETtableRate[indexTbl],1) ,MID(VAR_TICKETtable[indexTbl],6,1,VarTrimTemp) ,STOD(VarTrimTemp,VAR_TickettableItemNo[indexTbl]) ] [OTL(spTicketBinSet.16) ,ADD(indexTbl,1,indexTbl) ] ,XIC(spTicketBinActive.17) XIO(spTicketBinSet.17) [COP(spVAR_BINARRAY[17],VAR_TICKETtable[indexTbl],1) ,COP(spBinGateRates[17],VAR_TICKETtableRate[indexTbl],1) ,MID(VAR_TICKETtable[indexTbl],6,1,VarTrimTemp) ,STOD(VarTrimTemp,VAR_TickettableItemNo[indexTbl]) ] [OTL(spTicketBinSet.17) ,ADD(indexTbl,1,indexTbl) ] ,XIC(spTicketBinActive.21) XIO(spTicketBinSet.21) [COP(spVAR_BINARRAY[21],VAR_TICKETtable[indexTbl],1) ,COP(spBinGateRates[21],VAR_TICKETtableRate[indexTbl],1) ,MID(VAR_TICKETtable[indexTbl],6,1,VarTrimTemp) ,STOD(VarTrimTemp,VAR_TickettableItemNo[indexTbl]) ] [OTL(spTicketBinSet.21) ,ADD(indexTbl,1,indexTbl) ] ,XIC(spTicketBinActive.22) XIO(spTicketBinSet.22) [COP(spVAR_BINARRAY[22],VAR_TICKETtable[indexTbl],1) ,COP(spBinGateRates[22],VAR_TICKETtableRate[indexTbl],1) ,MID(VAR_TICKETtable[indexTbl],6,1,VarTrimTemp) ,STOD(VarTrimTemp,VAR_TickettableItemNo[indexTbl]) ] [OTL(spTicketBinSet.22) ,ADD(indexTbl,1,indexTbl) ] ,XIC(spTicketBinActive.23) XIO(spTicketBinSet.23) [COP(spVAR_BINARRAY[23],VAR_TICKETtable[indexTbl],1) ,COP(spBinGateRates[23],VAR_TICKETtableRate[indexTbl],1) ,MID(VAR_TICKETtable[indexTbl],6,1,VarTrimTemp) ,STOD(VarTrimTemp,VAR_TickettableItemNo[indexTbl]) ] [OTL(spTicketBinSet.23) ,ADD(indexTbl,1,indexTbl) ] ,XIC(spTicketBinActive.24) XIO(spTicketBinSet.24) [COP(spVAR_BINARRAY[24],VAR_TICKETtable[indexTbl],1) ,COP(spBinGateRates[24],VAR_TICKETtableRate[indexTbl],1) ,MID(VAR_TICKETtable[indexTbl],6,1,VarTrimTemp) ,STOD(VarTrimTemp,VAR_TickettableItemNo[indexTbl]) ] [OTL(spTicketBinSet.24) ,ADD(indexTbl,1,indexTbl) ] ,XIC(spTicketBinActive.25) XIO(spTicketBinSet.25) [COP(spVAR_BINARRAY[25],VAR_TICKETtable[indexTbl],1) ,COP(spBinGateRates[25],VAR_TICKETtableRate[indexTbl],1) ,MID(VAR_TICKETtable[indexTbl],6,1,VarTrimTemp) ,STOD(VarTrimTemp,VAR_TickettableItemNo[indexTbl]) ] [OTL(spTicketBinSet.25) ,ADD(indexTbl,1,indexTbl) ] ,XIC(spTicketBinActive.26) XIO(spTicketBinSet.26) [COP(spVAR_BINARRAY[26],VAR_TICKETtable[indexTbl],1) ,COP(spBinGateRates[26],VAR_TICKETtableRate[indexTbl],1) ,MID(VAR_TICKETtable[indexTbl],6,1,VarTrimTemp) ,STOD(VarTrimTemp,VAR_TickettableItemNo[indexTbl]) ] [OTL(spTicketBinSet.26) ,ADD(indexTbl,1,indexTbl) ] ];
